(* IEC 61131-3 sources: Gen-AI/docs/member2_validation/codesys_release_v1.1/C00_good, 1 file *)

(* ---- source.st ---- *)
FUNCTION_BLOCK FB_AgentProbeGood
VAR_INPUT
 x : BOOL;
END_VAR
VAR_OUTPUT
 y : BOOL;
END_VAR
y := x;
END_FUNCTION_BLOCK
